(* IEC 61131-3 sources: test/Network, 1 file *)

(* ---- ConfigObjects.st ---- *)
FUNCTION GLOBAL TAB TASK_CONF
_K_TASK, _K_REAL,
_K_END_VAR,

_K_TASK, _K_CYCLIC,
_K_END_VAR,

_K_TASK, _K_BACKGROUND,
_K_END_VAR,

_K_END_CONF
END_FUNCTION

FUNCTION GLOBAL TAB IPR_CONF
_K_IPR
	0$UINT,
_K_END_VAR,
_K_END_CONF
END_FUNCTION

FUNCTION GLOBAL TAB CONFIG_TABLES
00157$UINT,
0$UINT, 0, 11, "_ALARMDISPLAY",
0$UINT, 0, 1, "_BIT32",
0$UINT, 0, 1, "_BIT32RAM",
0$UINT, 0, 4, "_CAN",
0$UINT, 1, 10, "_CANLIB",
0$UINT, 1, 20, "_FILESYS",
0$UINT, 0, 15, "_GLOBAL",
0$UINT, 0, 1, "_HOTALARM",
0$UINT, 0, 5, "_LANGUAGESELECTION",
0$UINT, 0, 2, "_LIMITMAX",
0$UINT, 0, 2, "_LIMITMIN",
0$UINT, 0, 128, "_LSE",
0$UINT, 1, 1, "_MULTITASK",
0$UINT, 0, 3, "_MYIO",
0$UINT, 0, 5, "_OSKERNEL",
0$UINT, 0, 6, "_OSZILSE",
0$UINT, 0, 0, "_OSZILSEBACKGROUND",
0$UINT, 0, 1, "_RADIO32",
0$UINT, 0, 1, "_RADIO32RAM",
0$UINT, 0, 3, "_SCREEN",
0$UINT, 0, 15, "_SCROLLAREA",
0$UINT, 0, 8, "_SCROLLAREA2",
0$UINT, 1, 34, "_SERLIB",
0$UINT, 0, 0, "_STDLIB",
0$UINT, 0, 10, "_SYSDATETIME",
0$UINT, 0, 0, "_SYSDATETIME2",
0$UINT, 1, 1, "_TASKOBJECTCONTROL",
0$UINT, 1, 1, "_TOOLCAT",
0$UINT, 0, 1, "_XACCESS",
0$UINT, 1, 16, "AI040",
0$UINT, 1, 20, "AI043",
0$UINT, 1, 8, "AI046",
0$UINT, 1, 18, "AI084",
0$UINT, 1, 21, "ASCII_BIN",
0$UINT, 1, 26, "BUSINTERFACESDIAS",
0$UINT, 2, 1, "BUSINTERFACESDIASINTERNAL",
0$UINT, 1, 1, "CP112_IOS",
0$UINT, 0, 4, "CRITICALSECTION",
0$UINT, 0, 2, "DATASERVICECLIENT",
0$UINT, 2, 33, "DIASMASTER",
0$UINT, 1, 83, "DIASMASTERC",
0$UINT, 2, 25, "DIASMASTERMAIN",
0$UINT, 1, 0, "DIASMASTERPOSTSCAN",
0$UINT, 1, 14, "DM161",
0$UINT, 1, 20, "DUPLICATEAI043",
0$UINT, 1, 11, "EEPROM",
0$UINT, 0, 10, "GETBROADCASTDATA",
0$UINT, 0, 1, "GRAPHIC",
0$UINT, 0, 1, "HMIASCIIBUFFER",
0$UINT, 0, 0, "HMIBASELIST",
0$UINT, 0, 2, "HMICANSENDRECEIVE",
0$UINT, 0, 2, "HMICHKBITLIST",
0$UINT, 0, 0, "HMICOLORMAP",
0$UINT, 0, 16, "HMICOMPORT",
0$UINT, 0, 14, "HMICOMPORTCAN",
0$UINT, 0, 4, "HMIFILE",
0$UINT, 0, 2, "HMIFONT35",
0$UINT, 0, 3, "HMIFONTLIST",
0$UINT, 0, 2, "HMIFUNCTIONLIST",
0$UINT, 0, 4, "HMIFUNCTIONLIST35",
0$UINT, 0, 4, "HMIIMAGE35",
0$UINT, 0, 3, "HMIIMAGELIST",
0$UINT, 0, 0, "HMIMAPFILE",
0$UINT, 0, 0, "HMIMEMCIRCLE",
0$UINT, 0, 0, "HMIMEMIMAGE",
0$UINT, 0, 0, "HMIMEMIO",
0$UINT, 0, 0, "HMIMEMLINE",
0$UINT, 0, 0, "HMIMEMRECTANGLE",
0$UINT, 0, 0, "HMIMEMTEXT",
0$UINT, 0, 0, "HMIMEMZORDER",
0$UINT, 0, 7, "HMIPROJECT35",
0$UINT, 0, 2, "HMIPROJECTLIST",
0$UINT, 0, 1, "HMISCREEN",
0$UINT, 0, 2, "HMISETUPLIST",
0$UINT, 0, 3, "HMISETUPLIST35",
0$UINT, 0, 3, "HMISHEMELIST",
0$UINT, 0, 4, "HMISHEMELIST35",
0$UINT, 0, 5, "HMISTATEBIT35",
0$UINT, 0, 2, "HMISTRLIB",
0$UINT, 0, 0, "HMIT9CONFIG35",
0$UINT, 0, 4, "HMITEXTLIST",
0$UINT, 0, 3, "HMITEXTLIST35",
0$UINT, 0, 0, "HMITEXTLIST35MANAGER",
0$UINT, 0, 0, "HMIUNIBUFFER",
0$UINT, 0, 2, "HMIUNITLIST",
0$UINT, 0, 2, "HMIUTILS",
0$UINT, 0, 1, "HMIVARINFOLIST",
0$UINT, 0, 17, "HMIVARLIST",
0$UINT, 0, 5, "HMIVARLIST35",
0$UINT, 1, 21, "HUB_BASE",
0$UINT, 2, 11, "HUB_BASE_ROOT",
0$UINT, 2, 36, "HWBASE",
0$UINT, 2, 56, "HWBASECDIAS",
0$UINT, 1, 0, "HWCLOGGING",
0$UINT, 5, 19, "HWCONTROL",
0$UINT, 1, 10, "HWCONTROLBASE",
0$UINT, 1, 0, "HWKVARSIZEFIFO",
0$UINT, 1, 0, "HWRTPOSTSCAN",
0$UINT, 1, 6, "I2CCDIAS",
0$UINT, 1, 32, "LSEEASY",
0$UINT, 1, 22, "MERKEREX",
0$UINT, 0, 0, "PUMPCONTROL",
0$UINT, 1, 3, "RAM",
0$UINT, 1, 17, "RAMEX",
0$UINT, 1, 9, "RAMFILE",
0$UINT, 1, 33, "SAFETYBASEFSOE",
0$UINT, 3, 19, "SAFETYCDIAS_BASE",
0$UINT, 2, 24, "SAFETYMANAGER",
0$UINT, 1, 4, "SAFETYUDP",
0$UINT, 1, 41, "SCP111",
0$UINT, 0, 0, "SDCICLASS",
0$UINT, 1, 8, "SDCIDEVICE",
0$UINT, 1, 60, "SDIASBASE",
0$UINT, 1, 10, "SDIASHUBBASE",
0$UINT, 1, 97, "SDIASMANAGER",
0$UINT, 2, 6, "SDIASPLC",
0$UINT, 1, 10, "SDIASSAFETYBASE",
0$UINT, 1, 33, "SDIASSAFETYMANAGERFSOE",
0$UINT, 1, 14, "SDIASSDCIMASTER",
0$UINT, 1, 12, "SDM081",
0$UINT, 2, 0, "SFC_ACTION_BASE",
0$UINT, 2, 0, "SFC_ACTIONINVOKER",
0$UINT, 1, 2, "SFC_CLIENT_SPLITTER_10",
0$UINT, 1, 3, "SFC_CLIENT_SPLITTER_2",
0$UINT, 1, 2, "SFC_CLIENT_SPLITTER_3",
0$UINT, 1, 2, "SFC_CLIENT_SPLITTER_4",
0$UINT, 1, 2, "SFC_CLIENT_SPLITTER_BASE",
0$UINT, 1, 1, "SFC_LOGIC_OR_10",
0$UINT, 1, 1, "SFC_LOGIC_OR_2",
0$UINT, 1, 1, "SFC_LOGIC_OR_3",
0$UINT, 1, 1, "SFC_LOGIC_OR_4",
0$UINT, 1, 6, "SFC_LOGIC_OR_BASE",
0$UINT, 2, 0, "SFC_NETWORK_BASE",
0$UINT, 1, 0, "SFC_PARALLEL_HANDLER_BASE",
0$UINT, 1, 0, "SFC_SORT",
0$UINT, 1, 1, "SFC_STEP_BASE",
0$UINT, 1, 0, "SFC_STEPINVOKER",
0$UINT, 1, 2, "SFC_TRANSITION_BASE",
0$UINT, 0, 0, "SFCCLASS",
0$UINT, 0, 0, "SFCCLASS_ACTION0",
0$UINT, 0, 0, "SFCCLASS_INITSTEP",
0$UINT, 0, 0, "SFCCLASS_INTERNALVARHOLDER",
0$UINT, 0, 0, "SFCCLASS_STEP0",
0$UINT, 0, 0, "SFCCLASS_TRANSITION0",
0$UINT, 0, 0, "SFCCLASS_TRANSITION1",
0$UINT, 0, 37, "SIGCLIB",
0$UINT, 1, 11, "STRING",
0$UINT, 1, 85, "STRINGINTERNAL",
0$UINT, 1, 21, "SYNCCALL",
0$UINT, 0, 1, "SYSTEM",
0$UINT, 2, 18, "VARAN_BASE",
0$UINT, 3, 4, "VARANMANAGER",
0$UINT, 2, 4, "VARANMANAGER_1",
0$UINT, 1, 25, "VARANMANAGER_BASE",
0$UINT, 1, 3, "VIRTUALBASEINIT",
0$UINT, 2, 11, "WATCHDOGDIAS",
0$UINT, 1, 1, "XXXBASE_IOS",
ONE_CFG$UINT, 0, 0, "ONE_HW_Network",
ONE_CFG$UINT, 0, 0, "ONE_LseEasyMain",
ONE_CFG$UINT, 0, 0, "ONE_LseEasySettings",
ONE_CFG$UINT, 0, 0, "ONE_Pump",
ONE_CFG$UINT, 1, 0, "ONE_STDAccessControlExtended",
ONE_CFG$UINT, 2, 0, "ONE_STDSettingsHMI",
TASK_CFG$UINT, 0, 0, "TASK_CONF",
IPR_CFG$UINT, 0, 0, "IPR_CONF",
PRJ_CFG$UINT, 0, 0, "Copy pump",
END_FUNCTION

#ifdef __LSLLDR_IOELEMENTS__
FUNCTION GLOBAL TAB _IO_ELEMENTS_TAB
0001$UINT, 0003$UINT,
"IO_Element1", "AI0431.AI2",
"IO_Element2", "SDM0811.Safe_Input1",
"IO_Element3", "SDM0811.Safe_Input2",
0003$UINT,
"IO_Element1", "pumpControl1.ActFillLevel",
"IO_Element2", "pumpControl1.test2",
"IO_Element3", "pumpControl1.test1",
END_FUNCTION
#endif //__LSLLDR_IOELEMENTS__

FUNCTION GLOBAL TAB CH_REDIRECT_EMB_TAB
0000$UINT,
00019$UINT,
"AI040;SERIALNO", "\SERIALNOSTR.DATA",
"AI043;SERIALNO", "\SERIALNOSTR.DATA",
"AI046;SERIALNO", "\SERIALNOSTR.DATA",
"AI084;SERIALNO", "\SERIALNOSTR.DATA",
"BUSINTERFACESDIAS;SERIALNO", "\SERIALNOSTR.DATA",
"DM161;SERIALNO", "\SERIALNOSTR.DATA",
"DUPLICATEAI043;SERIALNO", "\SERIALNOSTR.DATA",
"HWBASECDIAS;SERIALNO", "\SERIALNOSTR.DATA",
"SAFETYCDIAS_BASE;SERIALNO", "\SERIALNOSTR.DATA",
"SCP111;DESIGNERPRJNAME", "\SDIASSAFETYMANAGERFSOE1\PROJECTNAMESTR.DATA",
"SCP111;DESIGNERPRJREV", "\SDIASSAFETYMANAGERFSOE1\PROJECTREVISIONSTR.DATA",
"SCP111;SERIALNO", "\SERIALNOSTR.DATA",
"SDIASBASE;SERIALNO", "\SERIALNOSTR.DATA",
"SDIASSAFETYBASE;SERIALNO", "\SERIALNOSTR.DATA",
"SDIASSAFETYMANAGERFSOE;DESIGNERPRJNAME", "\PROJECTNAMESTR.DATA",
"SDIASSAFETYMANAGERFSOE;DESIGNERPRJREV", "\PROJECTREVISIONSTR.DATA",
"SDIASSDCIMASTER;SERIALNO", "\SERIALNOSTR.DATA",
"SDM081;SERIALNO", "\SERIALNOSTR.DATA",
"VARAN_BASE;SERIALNO", "\SERIALNOSTR.DATA",
END_FUNCTION
